// TIA Portal V20 export
// export: Created 2026-11-12T11:17:34.0535629Z, ExportSetting WithDefaults, DisplayName Totally Integrated Automation Portal, DisplayVersion V20, DisplayName TIA Portal Openness, DisplayVersion V20, DisplayName TIA Portal Teamcenter Gateway, DisplayVersion V20, DisplayName TIA Portal Version Control Interface, DisplayVersion V20, DisplayName STEP 7 Professional, DisplayVersion V20, DisplayName STEP 7 CFC, DisplayVersion V20, DisplayName STEP 7 Safety, DisplayVersion V20, DisplayName WinCC Basic/Comfort/Advanced, DisplayVersion V20, DisplayName SIMATIC Visualization Architect, DisplayVersion V20, DisplayName WinCC Professional, DisplayVersion V20, DisplayName SIMATIC Visualization Architect, DisplayVersion V20, DisplayName WinCC Unified, DisplayVersion V20, DisplayName SIMATIC Visualization Architect, DisplayVersion V20
TYPE "UDT_Entradas_Basico"
// stored: IsFailsafeCompliant false
   STRUCT
      Boton_marcha : Bool;   // Botón de marcha
      Boton_paro : Bool;   // Botón de paro (0 activado)
      Selector_modo : Bool;   // Selector Manual/Auto (0 - Manual / 1 - Auto)
      Boton_rearme : Bool;   // Botón de rearme
      Sensor_ind_bien_pos : Bool;   // Palet bien posicionado - Sensor inductivo 0 (Extremo derecho)
      Seta_emergencia : Bool;   // Seta de emergencia
      Sensor_palet_izq : Bool;   // Palet en extremo izquierdo
      Sensor_palet_dch : Bool;   // Palet en extremo derecho
   END_STRUCT;
END_TYPE
